ADAPTER ConveyorReq (* Adapter Interface *)
  (* Standard: 61499-1 *)
  (* Version 0.0, 7/2/2026 *)
  PACKAGE Main;
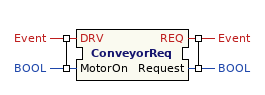
  EVENT_INPUT
    DRV WITH MotorOn;
  END_EVENT
  EVENT_OUTPUT
    REQ WITH Request;
  END_EVENT
  VAR_INPUT
    MotorOn : BOOL;
  END_VAR
  VAR_OUTPUT
    Request : BOOL;
  END_VAR
  SERVICE SOCKET/PLUG
    SEQUENCE request_confirm
      SOCKET.DRV(MotorOn) -> PLUG.DRV(MotorOn);
      PLUG.CNF(CNFD) -> SOCKET.CNF(CNFD);
    END_SEQUENCE
    SEQUENCE indication_response
      PLUG.REQ(Request) -> SOCKET.REQ(Request);
      SOCKET.RSP(RSPD) -> PLUG.RSP(RSPD);
    END_SEQUENCE
  END_SERVICE
END_ADAPTER
